    REGION SYSTEM 1
        IF "Screen_DB_1".Reset_All[2] AND
            (("HMI_Box_Connected_2" = 11 AND "KEY REMOTE/LOCAL L1 - CH1(1)") OR
            ("HMI_Box_Connected_2" = 12 AND "KEY REMOTE/LOCAL L2 - CH1(1)") OR
            ("HMI_Box_Connected_2" = 13 AND "KEY REMOTE/LOCAL L3 - CH1(1)") OR
            ("HMI_Box_Connected_2" = 14 AND "KEY REMOTE/LOCAL L4 - CH1(1)") OR
            ("HMI_Box_Connected_2" = 15 AND "KEY REMOTE/LOCAL L5 - CH1(1)") OR
            ("HMI_Box_Connected_2" = 16 AND "KEY REMOTE/LOCAL L6 - CH1(1)") OR
            ("HMI_Box_Connected_2" = 17 AND "KEY REMOTE/LOCAL L7 - CH1(1)") OR
            ("HMI_Box_Connected_2" = 18 AND "KEY REMOTE/LOCAL L8 - CH1(1)"))
        THEN
            "Errors_Profinet_1".%X4 :=
            "Errors_Profinet_1".%X5 :=
            "Errors_Profinet_1".%X6 :=
            "Errors_Profinet_1".%X7 :=
            "Errors_Profinet_1".%X8 :=
            "Errors_Profinet_1".%X9 :=
            "Errors_Profinet_1".%X11 :=
            "Errors_Profinet_1".%X12 :=
            "Errors_Profinet_1".%X14 :=
            "Errors_Profinet_1".%X15 :=
            "Errors_Profinet_2".%X0 :=
            "Errors_Profinet_2".%X1 :=
            "Errors_Profinet_2".%X2 :=
            "Errors_Profinet_2".%X3 :=
            "Errors_Profinet_2".%X4 :=
            "Errors_Profinet_2".%X5 :=
            "Errors_Profinet_2".%X6 :=
            "Errors_Profinet_2".%X7 :=
            "Errors_Profinet_2".%X8 :=
            "Errors_Profinet_2".%X9 :=
            "Errors_Profinet_2".%X10 :=
            "Errors_Profinet_2".%X11 :=
            "Errors_Profinet_2".%X12 :=
            "Errors_Profinet_2".%X13 :=
            "Errors_Profinet_2".%X14 :=
            "Errors_Profinet_2".%X15 :=
            "Errors_Profinet_3".%X0 :=
            "Errors_Profinet_3".%X8 :=
            "Errors_Profinet_5".%X5 :=
            "Errors_Profinet_7".%X2 :=
            "Errors_Profinet_8".%X7 :=
            "Errors_Profinet_9".%X7 :=
            "Errors_Profinet_9".%X8 :=
            "Errors_Profinet_9".%X9 :=
            "Errors_Profinet_9".%X10 :=
            "Errors_Profinet_9".%X11 :=
            "Errors_Profinet_9".%X12 :=
            "Errors_Profinet_9".%X13 :=

            "Erros_Supply_Feedback_1".%X0 :=
            "Erros_Supply_Feedback_1".%X10 :=
            "Erros_Supply_Feedback_1".%X11 :=
            "Erros_Supply_Feedback_1".%X12 :=
            "Erros_Supply_Feedback_1".%X15 :=

            "Erros_Supply_Feedback_3".%X0 :=
            "Erros_Supply_Feedback_3".%X1 :=
            "Erros_Supply_Feedback_3".%X2 :=
            "Erros_Supply_Feedback_3".%X3 :=

            "Estop_Error_Word_1".%X1 :=
            "Estop_Error_Word_1".%X2 :=
            "Estop_Error_Word_1".%X3 :=
            "Estop_Error_Word_1".%X4 :=
            "Estop_Error_Word_1".%X5 :=
            "Estop_Error_Word_1".%X6 :=
            "Estop_Error_Word_1".%X7 :=
            "Estop_Error_Word_1".%X8 :=
            "Estop_Error_Word_1".%X9 :=
            "Estop_Error_Word_1".%X10 :=
            "Estop_Error_Word_1".%X11 :=
            "Error_Word_Overhang".%X0 :=
            "Error_Word_Overhang".%X1 :=
            FALSE;

            "Sick Lector_Error code 1_2" :=
            "Erros_Supply_Feedback_2" :=
            "Linear Encoder_Device Errors 1" :=
            "Sick Lector_Error code 1" := 0;

            "Errors_Word_LightGuard_1".%X0 := FALSE;
            "Errors_Word_LightGuard_1".%X1 := FALSE;
        END_IF;
    END_REGION

    REGION SYSTEM 2
        IF "Screen_DB_1".Reset_All[2] AND
            (("HMI_Box_Connected_2" = 21 AND "KEY REMOTE/LOCAL L1 - CH1(2)") OR
            ("HMI_Box_Connected_2" = 22 AND "KEY REMOTE/LOCAL L2 - CH1(2)") OR
            ("HMI_Box_Connected_2" = 23 AND "KEY REMOTE/LOCAL L3 - CH1(2)") OR
            ("HMI_Box_Connected_2" = 24 AND "KEY REMOTE/LOCAL L4 - CH1(2)") OR
            ("HMI_Box_Connected_2" = 25 AND "KEY REMOTE/LOCAL L5 - CH1(2)") OR
            ("HMI_Box_Connected_2" = 26 AND "KEY REMOTE/LOCAL L6 - CH1(2)") OR
            ("HMI_Box_Connected_2" = 27 AND "KEY REMOTE/LOCAL L7 - CH1(2)") OR
            ("HMI_Box_Connected_2" = 28 AND "KEY REMOTE/LOCAL L8 - CH1(2)"))
        THEN
            "Errors_Profinet_3".%X3 :=
            "Errors_Profinet_3".%X6 :=
            "Errors_Profinet_3".%X7 :=
            "Errors_Profinet_3".%X8 :=
            "Errors_Profinet_3".%X9 :=
            "Errors_Profinet_3".%X10 :=
            "Errors_Profinet_3".%X11 :=
            "Errors_Profinet_3".%X12 :=
            "Errors_Profinet_3".%X13 :=
            "Errors_Profinet_3".%X14 :=
            "Errors_Profinet_4".%X0 :=
            "Errors_Profinet_4".%X1 :=
            "Errors_Profinet_4".%X2 :=
            "Errors_Profinet_4".%X3 :=
            "Errors_Profinet_4".%X4 :=
            "Errors_Profinet_4".%X5 :=
            "Errors_Profinet_4".%X6 :=
            "Errors_Profinet_4".%X7 :=
            "Errors_Profinet_4".%X8 :=
            "Errors_Profinet_4".%X9 :=
            "Errors_Profinet_4".%X10 :=
            "Errors_Profinet_4".%X11 :=
            "Errors_Profinet_4".%X12 :=
            "Errors_Profinet_4".%X13 :=
            "Errors_Profinet_4".%X14 :=
            "Errors_Profinet_5".%X5 :=
            "Errors_Profinet_7".%X2 :=
            "Errors_Profinet_8".%X7 :=
            "Errors_Profinet_9".%X7 :=
            "Errors_Profinet_9".%X8 :=
            "Errors_Profinet_9".%X9 :=
            "Errors_Profinet_9".%X10 :=
            "Errors_Profinet_9".%X14 :=
            "Errors_Profinet_9".%X15 :=
            "Errors_Profinet_10".%X0 :=
            "Errors_Profinet_10".%X1 :=

            "Erros_Supply_Feedback_1".%X1 :=
            "Erros_Supply_Feedback_1".%X10 :=
            "Erros_Supply_Feedback_1".%X11 :=
            "Erros_Supply_Feedback_1".%X12 :=
            "Erros_Supply_Feedback_1".%X15 :=

            "Erros_Supply_Feedback_3".%X4 :=
            "Erros_Supply_Feedback_3".%X5 :=
            "Erros_Supply_Feedback_3".%X6 :=
            "Erros_Supply_Feedback_3".%X7 :=
            "Erros_Supply_Feedback_3".%X8 :=
            "Erros_Supply_Feedback_3".%X9 :=
            "Erros_Supply_Feedback_3".%X10 :=
            "Erros_Supply_Feedback_3".%X11 :=
            "Erros_Supply_Feedback_3".%X12 :=
            "Erros_Supply_Feedback_3".%X13 :=
            "Erros_Supply_Feedback_3".%X14 :=
            "Erros_Supply_Feedback_3".%X15 :=
            "Erros_Supply_Feedback_4".%X0 :=
            "Erros_Supply_Feedback_4".%X1 :=
            "Erros_Supply_Feedback_4".%X2 :=
            "Erros_Supply_Feedback_4".%X3 :=
            "Erros_Supply_Feedback_4".%X4 :=
            "Erros_Supply_Feedback_4".%X5 :=
            "Erros_Supply_Feedback_4".%X6 :=
            "Erros_Supply_Feedback_4".%X7 :=

            "Estop_Error_Word_2".%X1 :=
            "Estop_Error_Word_2".%X2 :=
            "Estop_Error_Word_2".%X3 :=
            "Estop_Error_Word_2".%X4 :=
            "Estop_Error_Word_2".%X5 :=
            "Estop_Error_Word_2".%X6 :=
            "Estop_Error_Word_2".%X7 :=
            "Estop_Error_Word_2".%X8 :=
            "Estop_Error_Word_2".%X9 :=
            "Estop_Error_Word_2".%X10 :=
            "Estop_Error_Word_2".%X11 :=
            "Error_Word_Overhang".%X2 :=
            "Error_Word_Overhang".%X3 :=
            FALSE;

            "Sick Lector_Error code 2_2" :=
            "Linear Encoder_Device Errors 2" :=
            "Sick Lector_Error code 2" := 0;

            "Errors_Word_LightGuard_1".%X2 := FALSE;
            "Errors_Word_LightGuard_1".%X3 := FALSE;
        END_IF;
    END_REGION

    REGION SYSTEM 3
        IF "Screen_DB_1".Reset_All[2] AND
            (("HMI_Box_Connected_2" = 31 AND "KEY REMOTE/LOCAL L1 - CH1(3)") OR
            ("HMI_Box_Connected_2" = 32 AND "KEY REMOTE/LOCAL L2 - CH1(3)") OR
            ("HMI_Box_Connected_2" = 33 AND "KEY REMOTE/LOCAL L3 - CH1(3)") OR
            ("HMI_Box_Connected_2" = 34 AND "KEY REMOTE/LOCAL L4 - CH1(3)") OR
            ("HMI_Box_Connected_2" = 35 AND "KEY REMOTE/LOCAL L5 - CH1(3)") OR
            ("HMI_Box_Connected_2" = 36 AND "KEY REMOTE/LOCAL L6 - CH1(3)") OR
            ("HMI_Box_Connected_2" = 37 AND "KEY REMOTE/LOCAL L7 - CH1(3)") OR
            ("HMI_Box_Connected_2" = 38 AND "KEY REMOTE/LOCAL L8 - CH1(3)"))
        THEN
            "Errors_Profinet_3".%X8 :=
            "Errors_Profinet_5".%X0 :=
            "Errors_Profinet_5".%X2 :=
            "Errors_Profinet_5".%X3 :=
            "Errors_Profinet_5".%X4 :=
            "Errors_Profinet_5".%X5 :=
            "Errors_Profinet_5".%X6 :=
            "Errors_Profinet_5".%X7 :=
            "Errors_Profinet_5".%X8 :=
            "Errors_Profinet_5".%X9 :=
            "Errors_Profinet_5".%X10 :=
            "Errors_Profinet_5".%X12 :=
            "Errors_Profinet_5".%X13 :=
            "Errors_Profinet_5".%X14 :=
            "Errors_Profinet_5".%X15 :=
            "Errors_Profinet_6".%X0 :=
            "Errors_Profinet_6".%X1 :=
            "Errors_Profinet_6".%X2 :=
            "Errors_Profinet_6".%X3 :=
            "Errors_Profinet_6".%X4 :=
            "Errors_Profinet_6".%X5 :=
            "Errors_Profinet_6".%X6 :=
            "Errors_Profinet_6".%X7 :=
            "Errors_Profinet_6".%X8 :=
            "Errors_Profinet_6".%X9 :=
            "Errors_Profinet_6".%X10 :=
            "Errors_Profinet_6".%X11 :=
            "Errors_Profinet_7".%X2 :=
            "Errors_Profinet_8".%X7 :=
            "Errors_Profinet_9".%X7 :=
            "Errors_Profinet_9".%X8 :=
            "Errors_Profinet_9".%X9 :=
            "Errors_Profinet_9".%X10 :=
            "Errors_Profinet_10".%X2 :=
            "Errors_Profinet_10".%X3 :=
            "Errors_Profinet_10".%X4 :=
            "Errors_Profinet_10".%X5 :=

            "Erros_Supply_Feedback_4".%X8 :=
            "Erros_Supply_Feedback_4".%X9 :=
            "Erros_Supply_Feedback_4".%X10 :=
            "Erros_Supply_Feedback_4".%X11 :=
            "Erros_Supply_Feedback_4".%X12 :=
            "Erros_Supply_Feedback_4".%X13 :=
            "Erros_Supply_Feedback_4".%X14 :=
            "Erros_Supply_Feedback_4".%X15 :=
            "Erros_Supply_Feedback_5".%X0 :=
            "Erros_Supply_Feedback_5".%X1 :=
            "Erros_Supply_Feedback_5".%X2 :=
            "Erros_Supply_Feedback_5".%X3 :=
            "Erros_Supply_Feedback_5".%X4 :=
            "Erros_Supply_Feedback_5".%X5 :=
            "Erros_Supply_Feedback_5".%X6 :=
            "Erros_Supply_Feedback_5".%X7 :=
            "Erros_Supply_Feedback_5".%X8 :=
            "Erros_Supply_Feedback_5".%X9 :=
            "Erros_Supply_Feedback_5".%X10 :=
            "Erros_Supply_Feedback_5".%X11 :=

            "Estop_Error_Word_3".%X1 :=
            "Estop_Error_Word_3".%X2 :=
            "Estop_Error_Word_3".%X3 :=
            "Estop_Error_Word_3".%X4 :=
            "Estop_Error_Word_3".%X5 :=
            "Estop_Error_Word_3".%X6 :=
            "Estop_Error_Word_3".%X7 :=
            "Estop_Error_Word_3".%X8 :=
            "Estop_Error_Word_3".%X9 :=
            "Estop_Error_Word_3".%X10 :=
            "Estop_Error_Word_3".%X11 :=
            "Error_Word_Overhang".%X4 :=
            "Error_Word_Overhang".%X5 :=
            FALSE;

            "Sick Lector_Error code 3_2" :=
            "Linear Encoder_Device Errors 3" :=
            "Sick Lector_Error code 3" := 0;

            "Errors_Word_LightGuard_1".%X4 := FALSE;
            "Errors_Word_LightGuard_1".%X5 := FALSE;
        END_IF;
    END_REGION

    REGION SYSTEM 4
        IF "Screen_DB_1".Reset_All[2] AND
            (("HMI_Box_Connected_2" = 31 AND "KEY REMOTE/LOCAL L1 - CH1(3)") OR
            ("HMI_Box_Connected_2" = 32 AND "KEY REMOTE/LOCAL L2 - CH1(3)") OR
            ("HMI_Box_Connected_2" = 33 AND "KEY REMOTE/LOCAL L3 - CH1(3)") OR
            ("HMI_Box_Connected_2" = 34 AND "KEY REMOTE/LOCAL L4 - CH1(3)") OR
            ("HMI_Box_Connected_2" = 35 AND "KEY REMOTE/LOCAL L5 - CH1(3)") OR
            ("HMI_Box_Connected_2" = 36 AND "KEY REMOTE/LOCAL L6 - CH1(3)") OR
            ("HMI_Box_Connected_2" = 37 AND "KEY REMOTE/LOCAL L7 - CH1(3)") OR
            ("HMI_Box_Connected_2" = 38 AND "KEY REMOTE/LOCAL L8 - CH1(3)"))
        THEN
            "Errors_Profinet_3".%X8 :=
            "Errors_Profinet_5".%X5 :=
            "Errors_Profinet_6".%X13 :=
            "Errors_Profinet_6".%X15 :=
            "Errors_Profinet_7".%X0 :=
            "Errors_Profinet_7".%X1 :=
            "Errors_Profinet_7".%X2 :=
            "Errors_Profinet_7".%X3 :=
            "Errors_Profinet_7".%X4 :=
            "Errors_Profinet_7".%X5 :=
            "Errors_Profinet_7".%X6 :=
            "Errors_Profinet_7".%X7 :=
            "Errors_Profinet_7".%X8 :=
            "Errors_Profinet_7".%X9 :=
            "Errors_Profinet_7".%X10 :=
            "Errors_Profinet_7".%X11 :=
            "Errors_Profinet_7".%X12 :=
            "Errors_Profinet_7".%X13 :=
            "Errors_Profinet_7".%X14 :=
            "Errors_Profinet_7".%X15 :=
            "Errors_Profinet_8".%X0 :=
            "Errors_Profinet_8".%X7 :=
            "Errors_Profinet_9".%X7 :=
            "Errors_Profinet_9".%X8 :=
            "Errors_Profinet_9".%X9 :=
            "Errors_Profinet_9".%X10 :=
            "Errors_Profinet_10".%X6 :=
            "Errors_Profinet_10".%X7 :=
            "Errors_Profinet_10".%X8 :=
            "Errors_Profinet_10".%X9 :=

            "Erros_Supply_Feedback_5".%X12 :=
            "Erros_Supply_Feedback_5".%X13 :=
            "Erros_Supply_Feedback_5".%X14 :=
            "Erros_Supply_Feedback_5".%X15 :=
            "Erros_Supply_Feedback_6".%X0 :=
            "Erros_Supply_Feedback_6".%X1 :=
            "Erros_Supply_Feedback_6".%X2 :=
            "Erros_Supply_Feedback_6".%X3 :=
            "Erros_Supply_Feedback_6".%X4 :=
            "Erros_Supply_Feedback_6".%X5 :=
            "Erros_Supply_Feedback_6".%X6 :=
            "Erros_Supply_Feedback_6".%X7 :=

            "Estop_Error_Word_4".%X1 :=
            "Estop_Error_Word_4".%X2 :=
            "Estop_Error_Word_4".%X3 :=
            "Estop_Error_Word_4".%X4 :=
            "Estop_Error_Word_4".%X5 :=
            "Estop_Error_Word_4".%X6 :=
            "Estop_Error_Word_4".%X7 :=
            "Estop_Error_Word_4".%X8 :=
            "Estop_Error_Word_4".%X9 :=
            "Estop_Error_Word_4".%X10 :=
            "Error_Word_Overhang".%X6 :=
            "Error_Word_Overhang".%X7 :=
            FALSE;

            "Sick Lector_Error code 4_2" :=
            "Linear Encoder_Device Errors 4" :=
            "Sick Lector_Error code 4" := 0;
        END_IF;
    END_REGION

    REGION SYSTEM 5
        IF "Screen_DB_1".Reset_All[2] AND
            (("HMI_Box_Connected_2" = 51 AND "KEY REMOTE/LOCAL L1 - CH1(5)") OR
            ("HMI_Box_Connected_2" = 52 AND "KEY REMOTE/LOCAL L2 - CH1(5)") OR
            ("HMI_Box_Connected_2" = 53 AND "KEY REMOTE/LOCAL L3 - CH1(5)") OR
            ("HMI_Box_Connected_2" = 54 AND "KEY REMOTE/LOCAL L4 - CH1(5)") OR
            ("HMI_Box_Connected_2" = 55 AND "KEY REMOTE/LOCAL L5 - CH1(5)") OR
            ("HMI_Box_Connected_2" = 56 AND "KEY REMOTE/LOCAL L6 - CH1(5)") OR
            ("HMI_Box_Connected_2" = 57 AND "KEY REMOTE/LOCAL L7 - CH1(5)") OR
            ("HMI_Box_Connected_2" = 58 AND "KEY REMOTE/LOCAL L8 - CH1(5)"))
        THEN
            "Errors_Profinet_3".%X8 :=
            "Errors_Profinet_5".%X5 :=
            "Errors_Profinet_7".%X2 :=
            "Errors_Profinet_8".%X2 :=
            "Errors_Profinet_8".%X4 :=
            "Errors_Profinet_8".%X5 :=
            "Errors_Profinet_8".%X6 :=
            "Errors_Profinet_8".%X7 :=
            "Errors_Profinet_8".%X8 :=
            "Errors_Profinet_8".%X9 :=
            "Errors_Profinet_8".%X10 :=
            "Errors_Profinet_8".%X11 :=
            "Errors_Profinet_8".%X12 :=
            "Errors_Profinet_8".%X13 :=
            "Errors_Profinet_8".%X14 :=
            "Errors_Profinet_8".%X15 :=
            "Errors_Profinet_9".%X0 :=
            "Errors_Profinet_9".%X1 :=
            "Errors_Profinet_9".%X2 :=
            "Errors_Profinet_9".%X3 :=
            "Errors_Profinet_9".%X4 :=
            "Errors_Profinet_9".%X5 :=
            "Errors_Profinet_9".%X7 :=
            "Errors_Profinet_9".%X8 :=
            "Errors_Profinet_9".%X9 :=
            "Errors_Profinet_9".%X10 :=
            "Errors_Profinet_10".%X10 :=
            "Errors_Profinet_10".%X11 :=
            "Errors_Profinet_10".%X12 :=
            "Errors_Profinet_10".%X13 :=

            "Erros_Supply_Feedback_6".%X8 :=
            "Erros_Supply_Feedback_6".%X9 :=
            "Erros_Supply_Feedback_6".%X10 :=
            "Erros_Supply_Feedback_6".%X11 :=
            "Erros_Supply_Feedback_6".%X12 :=
            "Erros_Supply_Feedback_6".%X13 :=
            "Erros_Supply_Feedback_6".%X14 :=
            "Erros_Supply_Feedback_6".%X15 :=
            "Erros_Supply_Feedback_7".%X0 :=
            "Erros_Supply_Feedback_7".%X1 :=
            "Erros_Supply_Feedback_7".%X2 :=
            "Erros_Supply_Feedback_7".%X3 :=

            "Estop_Error_Word_5".%X1 :=
            "Estop_Error_Word_5".%X2 :=
            "Estop_Error_Word_5".%X3 :=
            "Estop_Error_Word_5".%X4 :=
            "Estop_Error_Word_5".%X5 :=
            "Estop_Error_Word_5".%X6 :=
            "Estop_Error_Word_5".%X7 :=
            "Estop_Error_Word_5".%X8 :=
            "Estop_Error_Word_5".%X9 :=
            "Estop_Error_Word_5".%X10 :=
            "Error_Word_Overhang".%X8 :=
            "Error_Word_Overhang".%X9 :=
            FALSE;

            "Sick Lector_Error code 5_2" :=
            "Linear Encoder_Device Errors 5" :=
            "Sick Lector_Error code 5" := 0;
        END_IF;
    END_REGION

END_REGION


END_FUNCTION